FUNCTION_BLOCK MOD_OwnerView (* Tells the block it sits in who occupies the module, and asks for it once at start. Technical: The module's occupation owner from its local channel; asks for the current value at INIT *)
  (* Standard: 61499-2 *)
  (* Version 0.1, 2026-09-28, Project contributors, AAU Smart Production Lab *)
  PACKAGE modlib;
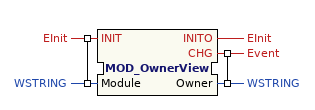
  EVENT_INPUT
    INIT : EInit WITH Module; (* Initialise, once at start-up (the INIT chain); takes the values given with it *)
  END_EVENT
  EVENT_OUTPUT
    INITO : EInit; (* Initialised: the next block of the INIT chain goes on *)
    CHG WITH Owner; (* The value changed *)
  END_EVENT
  VAR_INPUT
    Module : WSTRING; (* The module's name; its local channels are named after it (loc[<Module>/...]) *)
  END_VAR
  VAR_OUTPUT
    Owner : WSTRING; (* Session ID of the module's owner (empty: free) *)
  END_VAR
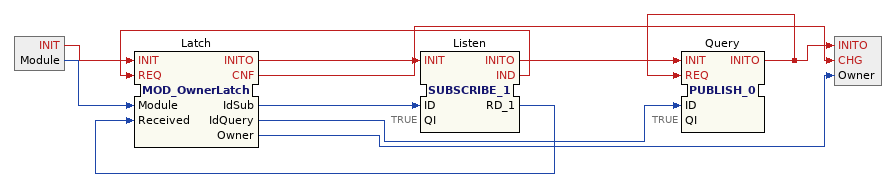
  FBS
    Latch : modlib::MOD_OwnerLatch; (* Keeps the last owner heard. *)
    Listen : iec61499::net::SUBSCRIBE_1(QI := TRUE); (* Listens to the owner channel. *)
    Query : iec61499::net::PUBLISH_0(QI := TRUE); (* Asks for the owner once at start. *)
  END_FBS
  EVENT_CONNECTIONS
    INIT TO Latch.INIT;
    Latch.INITO TO Listen.INIT;
    Listen.INITO TO Query.INIT;
    Query.INITO TO Query.REQ;
    Query.INITO TO INITO;
    Listen.IND TO Latch.REQ;
    Latch.CNF TO CHG;
  END_CONNECTIONS
  DATA_CONNECTIONS
    Module TO Latch.Module;
    Latch.IdSub TO Listen.ID;
    Latch.IdQuery TO Query.ID;
    Listen.RD_1 TO Latch.Received;
    Latch.Owner TO Owner;
  END_CONNECTIONS
END_FUNCTION_BLOCK
